Staubli VAL3: CalToolPos3.pgx

public program CalToolPos3(tool& x_tTool)
  local num ax1
  local num ax2
  local num ax3
  local num ay1
  local num ay2
  local num ay3
  local num az1
  local num az2
  local num az3
  local bool l_bStatus
  local pointRx l_p1
  local pointRx l_p2
  local pointRx l_p3
  local point l_pCenter
  local trsf l_trP1
  local trsf l_trP2
  local trsf l_trP3
  local num nx1
  local num nx2
  local num nx3
  local num ny1
  local num ny2
  local num ny3
  local num nz1
  local num nz2
  local num nz3
  local num ox1
  local num ox2
  local num ox3
  local num oy1
  local num oy2
  local num oy3
  local num oz1
  local num oz2
  local num oz3
  local num xf1
  local num xf2
  local num xf3
  local num yf1
  local num yf2
  local num yf3
  local num zf1
  local num zf2
  local num zf3
begin
  //3个带姿态的点求工具值XYZ
  l_trP1=db:pTeach1.trsf
  l_trP2=db:pTeach2.trsf
  l_trP3=db:pTeach3.trsf
  //
  //pTeach_3_1转成矩阵nTeach_3_1
  call matrix:Trsf2Matrix(l_trP1,nTeach_3_1)
  //pTeach_3_2转成矩阵nTeach_3_2
  call matrix:Trsf2Matrix(l_trP2,nTeach_3_2)
  //pTeach_3_3转成矩阵nTeach_3_3
  call matrix:Trsf2Matrix(l_trP3,nTeach_3_3)
  //
  //分解矩阵nTeach_3_1
  nx1=nTeach_3_1[0,0]
  ny1=nTeach_3_1[0,1]
  nz1=nTeach_3_1[0,2]
  ox1=nTeach_3_1[1,0]
  oy1=nTeach_3_1[1,1]
  oz1=nTeach_3_1[1,2]
  ax1=nTeach_3_1[2,0]
  ay1=nTeach_3_1[2,1]
  az1=nTeach_3_1[2,2]
  xf1=nTeach_3_1[3,0]
  yf1=nTeach_3_1[3,1]
  zf1=nTeach_3_1[3,2]
  //
  //分解矩阵nTeach_3_2
  nx2=nTeach_3_2[0,0]
  ny2=nTeach_3_2[0,1]
  nz2=nTeach_3_2[0,2]
  ox2=nTeach_3_2[1,0]
  oy2=nTeach_3_2[1,1]
  oz2=nTeach_3_2[1,2]
  ax2=nTeach_3_2[2,0]
  ay2=nTeach_3_2[2,1]
  az2=nTeach_3_2[2,2]
  xf2=nTeach_3_2[3,0]
  yf2=nTeach_3_2[3,1]
  zf2=nTeach_3_2[3,2]
  //
  //分解矩阵nTeach_3_3
  nx3=nTeach_3_3[0,0]
  ny3=nTeach_3_3[0,1]
  nz3=nTeach_3_3[0,2]
  ox3=nTeach_3_3[1,0]
  oy3=nTeach_3_3[1,1]
  oz3=nTeach_3_3[1,2]
  ax3=nTeach_3_3[2,0]
  ay3=nTeach_3_3[2,1]
  az3=nTeach_3_3[2,2]
  xf3=nTeach_3_3[3,0]
  yf3=nTeach_3_3[3,1]
  zf3=nTeach_3_3[3,2]
  //
  //***************************************************************************************
  //  │nx1-nx2 , ox1-ox2 , ax1-ax2 ,   0  │   │1 , 0 , 0, Tx│   │1 , 0 , 0, xf2-xf1│
  //  │ny2-ny3 , oy2-oy3 , ay2-ay3 ,   0  │ * │0 , 1 , 0, Ty│ = │0 , 1 , 0, yf3-yf2│
  //  │nz1-nz3 , oz1-oz3 , az1-az3 ,   0  │   │0 , 0 , 1, Tz│   │0 , 0 , 1, zf3-zf1│
  //  │   0    ,    0    ,    0    ,   1  │   │0 , 0 , 0,  1│   │0 , 0 , 0,    1   │
  //***************************************************************************************
  //构造矩阵nMatrix1
  nMatrix1[0,0]=nx1-nx2
  nMatrix1[0,1]=ny2-ny3
  nMatrix1[0,2]=nz1-nz3
  nMatrix1[0,3]=0
  nMatrix1[1,0]=ox1-ox2
  nMatrix1[1,1]=oy2-oy3
  nMatrix1[1,2]=oz1-oz3
  nMatrix1[1,3]=0
  nMatrix1[2,0]=ax1-ax2
  nMatrix1[2,1]=ay2-ay3
  nMatrix1[2,2]=az1-az3
  nMatrix1[2,3]=0
  nMatrix1[3,0]=0
  nMatrix1[3,1]=0
  nMatrix1[3,2]=0
  nMatrix1[3,3]=1

  //构造矩阵nMatrix2
  nMatrix2[0,0]=1
  nMatrix2[0,1]=0
  nMatrix2[0,2]=0
  nMatrix2[0,3]=0

  nMatrix2[1,0]=0
  nMatrix2[1,1]=1
  nMatrix2[1,2]=0
  nMatrix2[1,3]=0

  nMatrix2[2,0]=0
  nMatrix2[2,1]=0
  nMatrix2[2,2]=1
  nMatrix2[2,3]=0

  nMatrix2[3,0]=xf2-xf1
  nMatrix2[3,1]=yf3-yf2
  nMatrix2[3,2]=zf3-zf1
  nMatrix2[3,3]=1
  //***************************************************************************************
  call matrix:InverseMatrix(nMatrix1,nInverseMatrix1,l_bStatus)
  if l_bStatus==false
    //如果nMatrix1不可逆则需重新示教点
    call db:hmiAlert("DeviationIsTooLarge","warning")
  else
    call matrix:MutliMatrix(nInverseMatrix1,nMatrix2,nMatrix3)

    x_tTool.trsf.x=nMatrix3[3,0]
    x_tTool.trsf.y=nMatrix3[3,1]
    x_tTool.trsf.z=nMatrix3[3,2]
    x_tTool.trsf.rx=0
    x_tTool.trsf.ry=0
    x_tTool.trsf.rz=0
  endIf
  //定义中心点xyz
  l_pCenter.trsf=l_p1.trsf*x_tTool.trsf
  //定义中心点RxRyRz
  if db:sMounting=="Floor"
    l_pCenter.trsf.rx=0
    l_pCenter.trsf.ry=180
    l_pCenter.trsf.rz=0
  elseIf db:sMounting=="Ceiling"
    l_pCenter.trsf.rx=0
    l_pCenter.trsf.ry=0
    l_pCenter.trsf.rz=0
  endIf
  x_tTool.trsf=!l_p1.trsf*l_pCenter.trsf
  call db:hmiAlert("SaveInTool1","info")
end
